// TIA Portal V21 export
// export: Created 2026-08-21T20:18:51.7692183Z, ExportSetting None, DisplayName Totally Integrated Automation Portal, DisplayVersion V21, DisplayName STEP 7 Professional, DisplayVersion V21, DisplayName STEP 7 Safety, DisplayVersion V21, DisplayName Tech WebApplication, DisplayVersion V21, DisplayName WinCC Basic/Comfort/Advanced, DisplayVersion V21, DisplayName WinCC Professional, DisplayVersion V21, DisplayName WinCC Unified, DisplayVersion V21
DATA_BLOCK "FIT100_Type"   // DB2
// stored: InstanceOfName MTPAnaMon_Type1, InstanceOfType FB
"MTPAnaMon_Type1"
   // VAR_INPUT
   //    PV { ExternalAccessible := 'False'; ExternalVisible := 'False'; ExternalWritable := 'False'} : Word;
   //    PV_QB { ExternalAccessible := 'False'; ExternalVisible := 'False'; ExternalWritable := 'False'} : Bool;
   //    PV_Unit { ExternalAccessible := 'False'; ExternalVisible := 'False'; ExternalWritable := 'False'} : Int;
   //    PV_AH_En { ExternalAccessible := 'False'; ExternalVisible := 'False'; ExternalWritable := 'False'} : Bool := false;
   //    PV_WH_En { ExternalAccessible := 'False'; ExternalVisible := 'False'; ExternalWritable := 'False'} : Bool := false;
   //    PV_TH_En { ExternalAccessible := 'False'; ExternalVisible := 'False'; ExternalWritable := 'False'} : Bool;
   //    PV_TL_En { ExternalAccessible := 'False'; ExternalVisible := 'False'; ExternalWritable := 'False'} : Bool;
   //    PV_WL_En { ExternalAccessible := 'False'; ExternalVisible := 'False'; ExternalWritable := 'False'} : Bool := false;
   //    PV_AL_En { ExternalAccessible := 'False'; ExternalVisible := 'False'; ExternalWritable := 'False'} : Bool := false;
   // END_VAR
   // VAR_OUTPUT
   //    to_Indicate { ExternalAccessible := 'False'; ExternalVisible := 'False'; ExternalWritable := 'False'} : "StruCm";
   // END_VAR
   // VAR
   //    AnIn_IDB { ExternalAccessible := 'False'; ExternalVisible := 'False'; ExternalWritable := 'False'} : "AnIn";
   //    MonAnL_IDB : "MonAnL";
   //    MTPAnaMon_IDB { ExternalVisible := 'False'; S7_SetPoint := 'True'} : "MTPAnaMon";
   // END_VAR
BEGIN
   AnIn_IDB.Scale.High := 32.0;
   MonAnL_IDB.PV_AH_Lim := 40.0;
   MonAnL_IDB.PV_WH_Lim := 39.0;
   MonAnL_IDB.PV_TH_Lim := 38.0;
   MonAnL_IDB.PV_TL_Lim := 1.5;
   MonAnL_IDB.PV_WL_Lim := 1.0;
   MonAnL_IDB.PV_AL_Lim := 0.5;
   MonAnL_IDB.PV_AH_En := false;
   MonAnL_IDB.PV_WH_En := false;
   MonAnL_IDB.PV_WL_En := false;
   MonAnL_IDB.PV_AL_En := false;
   MonAnL_IDB.GradHUpEn := false;
   MonAnL_IDB.GradHDnEn := false;
END_DATA_BLOCK
